(* IEC 61131-3 sources: plc-st-coding-agent/progress/evidence/f14_v13_self_20261113/jobs/diagnostic_deepseek-v4pro, 15 files *)

(* ---- public-easy-01.candidate_01.st ---- *)
(* ENGINEERING_CONTRACT
Independent retained outputs, all reset by finishedButton:
- Pump_Motor: set when bottleSensor TRUE, holds until finishedButton.
- Filling_Valve: set when cleaningConfirmButton TRUE, holds until finishedButton.
- Capping_Machine: set when fillingConfirmButton TRUE, holds until finishedButton.
- Packing_Machine: set when cappingConfirmButton TRUE, holds until finishedButton.
- Completion_Light: set when packingConfirmButton TRUE, reset by finishedButton.
Same-scan priority: finishedButton reset first, then trigger evaluations.
*)
(* CONTRACT_RULES [{"kind":"hold_until_reset","output":"Pump_Motor","set_input":"bottleSensor","reset_input":"finishedButton"},{"kind":"hold_until_reset","output":"Filling_Valve","set_input":"cleaningConfirmButton","reset_input":"finishedButton"},{"kind":"hold_until_reset","output":"Capping_Machine","set_input":"fillingConfirmButton","reset_input":"finishedButton"},{"kind":"hold_until_reset","output":"Packing_Machine","set_input":"cappingConfirmButton","reset_input":"finishedButton"},{"kind":"hold_until_reset","output":"Completion_Light","set_input":"packingConfirmButton","reset_input":"finishedButton"}] *)

FUNCTION_BLOCK FillingLineControl
VAR_INPUT
    bottleSensor : BOOL;
    cleaningConfirmButton : BOOL;
    fillingConfirmButton : BOOL;
    cappingConfirmButton : BOOL;
    packingConfirmButton : BOOL;
    finishedButton : BOOL;
END_VAR
VAR_OUTPUT
    Pump_Motor : BOOL;
    Filling_Valve : BOOL;
    Capping_Machine : BOOL;
    Packing_Machine : BOOL;
    Completion_Light : BOOL;
END_VAR
VAR
END_VAR

IF finishedButton THEN
    Pump_Motor := FALSE;
    Filling_Valve := FALSE;
    Capping_Machine := FALSE;
    Packing_Machine := FALSE;
    Completion_Light := FALSE;
ELSE
    IF bottleSensor THEN
        Pump_Motor := TRUE;
    END_IF;

    IF cleaningConfirmButton THEN
        Filling_Valve := TRUE;
    END_IF;

    IF fillingConfirmButton THEN
        Capping_Machine := TRUE;
    END_IF;

    IF cappingConfirmButton THEN
        Packing_Machine := TRUE;
    END_IF;

    IF packingConfirmButton THEN
        Completion_Light := TRUE;
    END_IF;
END_IF;

END_FUNCTION_BLOCK

(* ---- public-easy-01.candidate_02.st ---- *)
(* ENGINEERING_CONTRACT
Independent retained outputs, all reset by finishedButton:
- Pump_Motor: set when bottleSensor TRUE, holds until finishedButton.
- Filling_Valve: set when cleaningConfirmButton TRUE, holds until finishedButton.
- Capping_Machine: set when fillingConfirmButton TRUE, holds until finishedButton.
- Packing_Machine: set when cappingConfirmButton TRUE and Capping_Machine active, holds until finishedButton.
- Completion_Light: set when packingConfirmButton TRUE and Packing_Machine active, reset by finishedButton.
Same-scan priority: finishedButton reset first, then trigger evaluations.
*)
(* CONTRACT_RULES [{"kind":"hold_until_reset","output":"Pump_Motor","set_input":"bottleSensor","reset_input":"finishedButton"},{"kind":"hold_until_reset","output":"Filling_Valve","set_input":"cleaningConfirmButton","reset_input":"finishedButton"},{"kind":"hold_until_reset","output":"Capping_Machine","set_input":"fillingConfirmButton","reset_input":"finishedButton"}] *)

FUNCTION_BLOCK FillingLineControl
VAR_INPUT
    bottleSensor : BOOL;
    cleaningConfirmButton : BOOL;
    fillingConfirmButton : BOOL;
    cappingConfirmButton : BOOL;
    packingConfirmButton : BOOL;
    finishedButton : BOOL;
END_VAR
VAR_OUTPUT
    Pump_Motor : BOOL;
    Filling_Valve : BOOL;
    Capping_Machine : BOOL;
    Packing_Machine : BOOL;
    Completion_Light : BOOL;
END_VAR
VAR
END_VAR

IF finishedButton THEN
    Pump_Motor := FALSE;
    Filling_Valve := FALSE;
    Capping_Machine := FALSE;
    Packing_Machine := FALSE;
    Completion_Light := FALSE;
ELSE
    IF bottleSensor THEN
        Pump_Motor := TRUE;
    END_IF;

    IF cleaningConfirmButton THEN
        Filling_Valve := TRUE;
    END_IF;

    IF fillingConfirmButton THEN
        Capping_Machine := TRUE;
    END_IF;

    IF cappingConfirmButton AND Capping_Machine THEN
        Packing_Machine := TRUE;
    END_IF;

    IF packingConfirmButton AND Packing_Machine THEN
        Completion_Light := TRUE;
    END_IF;
END_IF;

END_FUNCTION_BLOCK

(* ---- public-easy-01.candidate_03.st ---- *)
(* ENGINEERING_CONTRACT
Independent retained outputs, all reset by finishedButton:
- Pump_Motor: set when bottleSensor TRUE, holds until finishedButton.
- Filling_Valve: set when cleaningConfirmButton TRUE, holds until finishedButton.
- Capping_Machine: set when fillingConfirmButton TRUE, holds until finishedButton.
- Packing_Machine: set when cappingConfirmButton TRUE and Capping_Machine active, holds until finishedButton.
- Completion_Light: set when packingConfirmButton TRUE and Packing_Machine active, reset by finishedButton.
Same-scan priority: finishedButton reset first, then trigger evaluations.
*)
(* CONTRACT_RULES [{"kind":"hold_until_reset","output":"Pump_Motor","set_input":"bottleSensor","reset_input":"finishedButton"},{"kind":"hold_until_reset","output":"Filling_Valve","set_input":"cleaningConfirmButton","reset_input":"finishedButton"},{"kind":"hold_until_reset","output":"Capping_Machine","set_input":"fillingConfirmButton","reset_input":"finishedButton"}] *)

FUNCTION_BLOCK FillingLineControl
VAR_INPUT
    bottleSensor : BOOL;
    cleaningConfirmButton : BOOL;
    fillingConfirmButton : BOOL;
    cappingConfirmButton : BOOL;
    packingConfirmButton : BOOL;
    finishedButton : BOOL;
END_VAR
VAR_OUTPUT
    Pump_Motor : BOOL;
    Filling_Valve : BOOL;
    Capping_Machine : BOOL;
    Packing_Machine : BOOL;
    Completion_Light : BOOL;
END_VAR
VAR
    local_PumpPrev : BOOL;
    local_FillingPrev : BOOL;
    local_CappingPrev : BOOL;
    local_PackingPrev : BOOL;
END_VAR

local_PumpPrev := Pump_Motor;
local_FillingPrev := Filling_Valve;
local_CappingPrev := Capping_Machine;
local_PackingPrev := Packing_Machine;

IF finishedButton THEN
    Pump_Motor := FALSE;
    Filling_Valve := FALSE;
    Capping_Machine := FALSE;
    Packing_Machine := FALSE;
    Completion_Light := FALSE;
ELSE
    IF bottleSensor THEN
        Pump_Motor := TRUE;
    END_IF;

    IF cleaningConfirmButton AND local_PumpPrev THEN
        Filling_Valve := TRUE;
    END_IF;

    IF fillingConfirmButton AND local_FillingPrev THEN
        Capping_Machine := TRUE;
    END_IF;

    IF cappingConfirmButton AND local_CappingPrev THEN
        Packing_Machine := TRUE;
    END_IF;

    IF packingConfirmButton AND local_PackingPrev THEN
        Completion_Light := TRUE;
    END_IF;
END_IF;

END_FUNCTION_BLOCK

(* ---- public-easy-01.patch_base_01.st ---- *)
(* ENGINEERING_CONTRACT
Outputs by state (state is persistent across scans):
- Pump_Motor: ON in CLEANING; starts when bottleSensor TRUE from IDLE; OFF on cleaningConfirmButton. Retained while CLEANING, even if bottleSensor falls (PUB001/PUB002).
- Filling_Valve: ON in FILLING; starts on cleaningConfirmButton in CLEANING; OFF on fillingConfirmButton (PUB002/PUB003).
- Capping_Machine: ON in CAPPING; starts on fillingConfirmButton in FILLING; OFF on cappingConfirmButton (PUB003/PUB004).
- Packing_Machine: ON in PACKING; starts on cappingConfirmButton in CAPPING; OFF on packingConfirmButton (PUB004/PUB005).
- Completion_Light: ON in COMPLETE; starts on packingConfirmButton in PACKING; reset by finishedButton (PUB005/PUB006/PUB007).
Same-scan priority: one state transition per call via ELSIF chain; outputs are assigned after transition using final state.
Buttons are treated as level-sensitive; pulse width/protocol unspecified.
*)
(* CONTRACT_RULES [] *)

FUNCTION_BLOCK FillingLineControl
VAR_INPUT
    bottleSensor: BOOL;
    cleaningConfirmButton: BOOL;
    fillingConfirmButton: BOOL;
    cappingConfirmButton: BOOL;
    packingConfirmButton: BOOL;
    finishedButton: BOOL;
END_VAR
VAR_OUTPUT
    Pump_Motor: BOOL;
    Filling_Valve: BOOL;
    Capping_Machine: BOOL;
    Packing_Machine: BOOL;
    Completion_Light: BOOL;
END_VAR
VAR
    step: INT := 0; (* 0=IDLE, 1=CLEANING, 2=FILLING, 3=CAPPING, 4=PACKING, 5=COMPLETE *)
    bottleTrig: R_TRIG;
END_VAR

(* State transitions: at most one per scan *)
bottleTrig(CLK := bottleSensor);

IF step = 0 THEN
    IF bottleTrig.Q THEN
        step := 1;
    END_IF;
ELSIF step = 1 THEN
    IF cleaningConfirmButton THEN
        step := 2;
    END_IF;
ELSIF step = 2 THEN
    IF fillingConfirmButton THEN
        step := 3;
    END_IF;
ELSIF step = 3 THEN
    IF cappingConfirmButton THEN
        step := 4;
    END_IF;
ELSIF step = 4 THEN
    IF packingConfirmButton THEN
        step := 5;
    END_IF;
ELSIF step = 5 THEN
    IF finishedButton THEN
        step := 0;
    END_IF;
END_IF;

(* Output mapping based on final state *)
CASE step OF
    0:
        Pump_Motor := FALSE;
        Filling_Valve := FALSE;
        Capping_Machine := FALSE;
        Packing_Machine := FALSE;
        Completion_Light := FALSE;

    1:
        Pump_Motor := TRUE;
        Filling_Valve := FALSE;
        Capping_Machine := FALSE;
        Packing_Machine := FALSE;
        Completion_Light := FALSE;

    2:
        Pump_Motor := FALSE;
        Filling_Valve := TRUE;
        Capping_Machine := FALSE;
        Packing_Machine := FALSE;
        Completion_Light := FALSE;

    3:
        Pump_Motor := FALSE;
        Filling_Valve := FALSE;
        Capping_Machine := TRUE;
        Packing_Machine := FALSE;
        Completion_Light := FALSE;

    4:
        Pump_Motor := FALSE;
        Filling_Valve := FALSE;
        Capping_Machine := FALSE;
        Packing_Machine := TRUE;
        Completion_Light := FALSE;

    5:
        Pump_Motor := FALSE;
        Filling_Valve := FALSE;
        Capping_Machine := FALSE;
        Packing_Machine := FALSE;
        Completion_Light := TRUE;

    ELSE
        Pump_Motor := FALSE;
        Filling_Valve := FALSE;
        Capping_Machine := FALSE;
        Packing_Machine := FALSE;
        Completion_Light := FALSE;
END_CASE;

END_FUNCTION_BLOCK

(* ---- public-easy-01.patch_base_02.st ---- *)
(* ENGINEERING_CONTRACT
Independent retained outputs, all reset by finishedButton:
- Pump_Motor: set when bottleSensor TRUE, holds until finishedButton.
- Filling_Valve: set when cleaningConfirmButton TRUE, holds until finishedButton.
- Capping_Machine: set when fillingConfirmButton TRUE, holds until finishedButton.
- Packing_Machine: set when cappingConfirmButton TRUE, holds until finishedButton.
- Completion_Light: set when packingConfirmButton TRUE, reset by finishedButton.
Same-scan priority: finishedButton reset first, then trigger evaluations.
*)
(* CONTRACT_RULES [{"kind":"hold_until_reset","output":"Pump_Motor","set_input":"bottleSensor","reset_input":"finishedButton"},{"kind":"hold_until_reset","output":"Filling_Valve","set_input":"cleaningConfirmButton","reset_input":"finishedButton"},{"kind":"hold_until_reset","output":"Capping_Machine","set_input":"fillingConfirmButton","reset_input":"finishedButton"},{"kind":"hold_until_reset","output":"Packing_Machine","set_input":"cappingConfirmButton","reset_input":"finishedButton"},{"kind":"hold_until_reset","output":"Completion_Light","set_input":"packingConfirmButton","reset_input":"finishedButton"}] *)

FUNCTION_BLOCK FillingLineControl
VAR_INPUT
    bottleSensor : BOOL;
    cleaningConfirmButton : BOOL;
    fillingConfirmButton : BOOL;
    cappingConfirmButton : BOOL;
    packingConfirmButton : BOOL;
    finishedButton : BOOL;
END_VAR
VAR_OUTPUT
    Pump_Motor : BOOL;
    Filling_Valve : BOOL;
    Capping_Machine : BOOL;
    Packing_Machine : BOOL;
    Completion_Light : BOOL;
END_VAR
VAR
END_VAR

IF finishedButton THEN
    Pump_Motor := FALSE;
    Filling_Valve := FALSE;
    Capping_Machine := FALSE;
    Packing_Machine := FALSE;
    Completion_Light := FALSE;
ELSE
    IF bottleSensor THEN
        Pump_Motor := TRUE;
    END_IF;

    IF cleaningConfirmButton THEN
        Filling_Valve := TRUE;
    END_IF;

    IF fillingConfirmButton THEN
        Capping_Machine := TRUE;
    END_IF;

    IF cappingConfirmButton THEN
        Packing_Machine := TRUE;
    END_IF;

    IF packingConfirmButton THEN
        Completion_Light := TRUE;
    END_IF;
END_IF;

END_FUNCTION_BLOCK

(* ---- public-easy-01.patch_base_03.st ---- *)
(* ENGINEERING_CONTRACT
Independent retained outputs, all reset by finishedButton:
- Pump_Motor: set when bottleSensor TRUE, holds until finishedButton.
- Filling_Valve: set when cleaningConfirmButton TRUE, holds until finishedButton.
- Capping_Machine: set when fillingConfirmButton TRUE, holds until finishedButton.
- Packing_Machine: set when cappingConfirmButton TRUE and Capping_Machine active, holds until finishedButton.
- Completion_Light: set when packingConfirmButton TRUE and Packing_Machine active, reset by finishedButton.
Same-scan priority: finishedButton reset first, then trigger evaluations.
*)
(* CONTRACT_RULES [{"kind":"hold_until_reset","output":"Pump_Motor","set_input":"bottleSensor","reset_input":"finishedButton"},{"kind":"hold_until_reset","output":"Filling_Valve","set_input":"cleaningConfirmButton","reset_input":"finishedButton"},{"kind":"hold_until_reset","output":"Capping_Machine","set_input":"fillingConfirmButton","reset_input":"finishedButton"}] *)

FUNCTION_BLOCK FillingLineControl
VAR_INPUT
    bottleSensor : BOOL;
    cleaningConfirmButton : BOOL;
    fillingConfirmButton : BOOL;
    cappingConfirmButton : BOOL;
    packingConfirmButton : BOOL;
    finishedButton : BOOL;
END_VAR
VAR_OUTPUT
    Pump_Motor : BOOL;
    Filling_Valve : BOOL;
    Capping_Machine : BOOL;
    Packing_Machine : BOOL;
    Completion_Light : BOOL;
END_VAR
VAR
END_VAR

IF finishedButton THEN
    Pump_Motor := FALSE;
    Filling_Valve := FALSE;
    Capping_Machine := FALSE;
    Packing_Machine := FALSE;
    Completion_Light := FALSE;
ELSE
    IF bottleSensor THEN
        Pump_Motor := TRUE;
    END_IF;

    IF cleaningConfirmButton THEN
        Filling_Valve := TRUE;
    END_IF;

    IF fillingConfirmButton THEN
        Capping_Machine := TRUE;
    END_IF;

    IF cappingConfirmButton AND Capping_Machine THEN
        Packing_Machine := TRUE;
    END_IF;

    IF packingConfirmButton AND Packing_Machine THEN
        Completion_Light := TRUE;
    END_IF;
END_IF;

END_FUNCTION_BLOCK

(* ---- public-easy-01.raw_candidate_01.st ---- *)
(* ENGINEERING_CONTRACT
Independent retained outputs, all reset by finishedButton:
- Pump_Motor: set when bottleSensor TRUE, holds until finishedButton.
- Filling_Valve: set when cleaningConfirmButton TRUE, holds until finishedButton.
- Capping_Machine: set when fillingConfirmButton TRUE, holds until finishedButton.
- Packing_Machine: set when cappingConfirmButton TRUE, holds until finishedButton.
- Completion_Light: set when packingConfirmButton TRUE, reset by finishedButton.
Same-scan priority: finishedButton reset first, then trigger evaluations.
*)
(* CONTRACT_RULES [{"kind":"hold_until_reset","output":"Pump_Motor","set_input":"bottleSensor","reset_input":"finishedButton"},{"kind":"hold_until_reset","output":"Filling_Valve","set_input":"cleaningConfirmButton","reset_input":"finishedButton"},{"kind":"hold_until_reset","output":"Capping_Machine","set_input":"fillingConfirmButton","reset_input":"finishedButton"},{"kind":"hold_until_reset","output":"Packing_Machine","set_input":"cappingConfirmButton","reset_input":"finishedButton"},{"kind":"hold_until_reset","output":"Completion_Light","set_input":"packingConfirmButton","reset_input":"finishedButton"}] *)

FUNCTION_BLOCK FillingLineControl
VAR_INPUT
    bottleSensor : BOOL;
    cleaningConfirmButton : BOOL;
    fillingConfirmButton : BOOL;
    cappingConfirmButton : BOOL;
    packingConfirmButton : BOOL;
    finishedButton : BOOL;
END_VAR
VAR_OUTPUT
    Pump_Motor : BOOL;
    Filling_Valve : BOOL;
    Capping_Machine : BOOL;
    Packing_Machine : BOOL;
    Completion_Light : BOOL;
END_VAR
VAR
END_VAR

IF finishedButton THEN
    Pump_Motor := FALSE;
    Filling_Valve := FALSE;
    Capping_Machine := FALSE;
    Packing_Machine := FALSE;
    Completion_Light := FALSE;
ELSE
    IF bottleSensor THEN
        Pump_Motor := TRUE;
    END_IF;

    IF cleaningConfirmButton THEN
        Filling_Valve := TRUE;
    END_IF;

    IF fillingConfirmButton THEN
        Capping_Machine := TRUE;
    END_IF;

    IF cappingConfirmButton THEN
        Packing_Machine := TRUE;
    END_IF;

    IF packingConfirmButton THEN
        Completion_Light := TRUE;
    END_IF;
END_IF;

END_FUNCTION_BLOCK

(* ---- public-easy-01.raw_candidate_02.st ---- *)
(* ENGINEERING_CONTRACT
Independent retained outputs, all reset by finishedButton:
- Pump_Motor: set when bottleSensor TRUE, holds until finishedButton.
- Filling_Valve: set when cleaningConfirmButton TRUE, holds until finishedButton.
- Capping_Machine: set when fillingConfirmButton TRUE, holds until finishedButton.
- Packing_Machine: set when cappingConfirmButton TRUE and Capping_Machine active, holds until finishedButton.
- Completion_Light: set when packingConfirmButton TRUE and Packing_Machine active, reset by finishedButton.
Same-scan priority: finishedButton reset first, then trigger evaluations.
*)
(* CONTRACT_RULES [{"kind":"hold_until_reset","output":"Pump_Motor","set_input":"bottleSensor","reset_input":"finishedButton"},{"kind":"hold_until_reset","output":"Filling_Valve","set_input":"cleaningConfirmButton","reset_input":"finishedButton"},{"kind":"hold_until_reset","output":"Capping_Machine","set_input":"fillingConfirmButton","reset_input":"finishedButton"}] *)

FUNCTION_BLOCK FillingLineControl
VAR_INPUT
    bottleSensor : BOOL;
    cleaningConfirmButton : BOOL;
    fillingConfirmButton : BOOL;
    cappingConfirmButton : BOOL;
    packingConfirmButton : BOOL;
    finishedButton : BOOL;
END_VAR
VAR_OUTPUT
    Pump_Motor : BOOL;
    Filling_Valve : BOOL;
    Capping_Machine : BOOL;
    Packing_Machine : BOOL;
    Completion_Light : BOOL;
END_VAR
VAR
END_VAR

IF finishedButton THEN
    Pump_Motor := FALSE;
    Filling_Valve := FALSE;
    Capping_Machine := FALSE;
    Packing_Machine := FALSE;
    Completion_Light := FALSE;
ELSE
    IF bottleSensor THEN
        Pump_Motor := TRUE;
    END_IF;

    IF cleaningConfirmButton THEN
        Filling_Valve := TRUE;
    END_IF;

    IF fillingConfirmButton THEN
        Capping_Machine := TRUE;
    END_IF;

    IF cappingConfirmButton AND Capping_Machine THEN
        Packing_Machine := TRUE;
    END_IF;

    IF packingConfirmButton AND Packing_Machine THEN
        Completion_Light := TRUE;
    END_IF;
END_IF;

END_FUNCTION_BLOCK

(* ---- public-easy-01.raw_candidate_03.st ---- *)
(* ENGINEERING_CONTRACT
Independent retained outputs, all reset by finishedButton:
- Pump_Motor: set when bottleSensor TRUE, holds until finishedButton.
- Filling_Valve: set when cleaningConfirmButton TRUE, holds until finishedButton.
- Capping_Machine: set when fillingConfirmButton TRUE, holds until finishedButton.
- Packing_Machine: set when cappingConfirmButton TRUE and Capping_Machine active, holds until finishedButton.
- Completion_Light: set when packingConfirmButton TRUE and Packing_Machine active, reset by finishedButton.
Same-scan priority: finishedButton reset first, then trigger evaluations.
*)
(* CONTRACT_RULES [{"kind":"hold_until_reset","output":"Pump_Motor","set_input":"bottleSensor","reset_input":"finishedButton"},{"kind":"hold_until_reset","output":"Filling_Valve","set_input":"cleaningConfirmButton","reset_input":"finishedButton"},{"kind":"hold_until_reset","output":"Capping_Machine","set_input":"fillingConfirmButton","reset_input":"finishedButton"}] *)

FUNCTION_BLOCK FillingLineControl
VAR_INPUT
    bottleSensor : BOOL;
    cleaningConfirmButton : BOOL;
    fillingConfirmButton : BOOL;
    cappingConfirmButton : BOOL;
    packingConfirmButton : BOOL;
    finishedButton : BOOL;
END_VAR
VAR_OUTPUT
    Pump_Motor : BOOL;
    Filling_Valve : BOOL;
    Capping_Machine : BOOL;
    Packing_Machine : BOOL;
    Completion_Light : BOOL;
END_VAR
VAR
    local_PumpPrev : BOOL;
    local_FillingPrev : BOOL;
    local_CappingPrev : BOOL;
    local_PackingPrev : BOOL;
END_VAR

local_PumpPrev := Pump_Motor;
local_FillingPrev := Filling_Valve;
local_CappingPrev := Capping_Machine;
local_PackingPrev := Packing_Machine;

IF finishedButton THEN
    Pump_Motor := FALSE;
    Filling_Valve := FALSE;
    Capping_Machine := FALSE;
    Packing_Machine := FALSE;
    Completion_Light := FALSE;
ELSE
    IF bottleSensor THEN
        Pump_Motor := TRUE;
    END_IF;

    IF cleaningConfirmButton AND local_PumpPrev THEN
        Filling_Valve := TRUE;
    END_IF;

    IF fillingConfirmButton AND local_FillingPrev THEN
        Capping_Machine := TRUE;
    END_IF;

    IF cappingConfirmButton AND local_CappingPrev THEN
        Packing_Machine := TRUE;
    END_IF;

    IF packingConfirmButton AND local_PackingPrev THEN
        Completion_Light := TRUE;
    END_IF;
END_IF;

END_FUNCTION_BLOCK

(* ---- public-hard-04.candidate_01.st ---- *)
(* ENGINEERING_CONTRACT
   elementCount DINT: retained process value; 0 after reset, +1 successful enqueue, -1 successful dequeue, held otherwise; range 0..capacity.
   status WORD: overwritten every invocation; 0 idle/reset/success, 16#8002 rejected full enqueue, 16#8001 rejected empty dequeue; reset priority sets 0.
   queue state: first invocation empty; reset priority clears head/tail/count; enqueue writes at tail, dequeue reads head; circular indices low..high.
   edge triggers: R_TRIG consumed every scan; reset priority ignores edge requests; simultaneous enqueue+dequeue unspecified -> no-op.
   units/boundaries: capacity positive DINT derived each scan from LOWER_BOUND/UPPER_BOUND of the supplied array; first element index may be nonzero.
*)
(* CONTRACT_RULES [] *)
FUNCTION_BLOCK FIFO
VAR_INPUT
    enqueue : BOOL;
    dequeue : BOOL;
    reset : BOOL;
END_VAR
VAR_OUTPUT
    elementCount : DINT;
    status : WORD;
END_VAR
VAR_IN_OUT
    item : VARIANT;
    buffer : VARIANT;
END_VAR
VAR
    local_rEnq : R_TRIG;
    local_rDeq : R_TRIG;
    local_enqEdge : BOOL;
    local_deqEdge : BOOL;

    local_low : DINT;
    local_high : DINT;
    local_capacity : DINT;
    local_count : DINT := 0;
    local_head : DINT := 0;
    local_tail : DINT := 0;
END_VAR

local_rEnq(CLK := enqueue);
local_enqEdge := local_rEnq.Q;
local_rDeq(CLK := dequeue);
local_deqEdge := local_rDeq.Q;

status := 16#0000;

local_low := LOWER_BOUND(buffer, 1);
local_high := UPPER_BOUND(buffer, 1);
local_capacity := local_high - local_low + 1;
IF local_capacity < 1 THEN
    local_capacity := 1;
END_IF;

IF local_count = 0 THEN
    local_head := local_low;
    local_tail := local_low;
END_IF;

IF reset THEN
    local_count := 0;
    local_head := local_low;
    local_tail := local_low;
    status := 16#0000;
ELSE
    IF local_enqEdge AND NOT local_deqEdge THEN
        IF local_count < local_capacity THEN
            buffer[local_tail] := item;
            local_tail := local_tail + 1;
            IF local_tail > local_high THEN
                local_tail := local_low;
            END_IF;
            local_count := local_count + 1;
            status := 16#0000;
        ELSE
            status := 16#8002;
        END_IF;
    ELSIF local_deqEdge AND NOT local_enqEdge THEN
        IF local_count > 0 THEN
            item := buffer[local_head];
            local_head := local_head + 1;
            IF local_head > local_high THEN
                local_head := local_low;
            END_IF;
            local_count := local_count - 1;
            status := 16#0000;
        ELSE
            status := 16#8001;
        END_IF;
    END_IF;
END_IF;

elementCount := local_count;

(* ---- public-hard-04.candidate_02.st ---- *)
(* ENGINEERING_CONTRACT
   elementCount DINT: retained process value; 0 after reset, +1 successful enqueue, -1 successful dequeue, held otherwise; range 0..capacity.
   status WORD: overwritten every invocation; 0 idle/reset/success, 16#8002 rejected full enqueue, 16#8001 rejected empty dequeue; reset priority sets 0.
   queue state: first invocation empty; reset priority clears head/tail/count; enqueue writes at tail, dequeue reads head; circular indices low..high.
   edge triggers: R_TRIG consumed every scan; reset priority ignores edge requests; simultaneous enqueue+dequeue unspecified -> no-op.
   units/boundaries: capacity positive DINT derived each scan from LOWER_BOUND/UPPER_BOUND of the supplied array; first element index may be nonzero.
*)
(* CONTRACT_RULES [] *)
FUNCTION_BLOCK FIFO
VAR_INPUT
    enqueue : BOOL;
    dequeue : BOOL;
    reset : BOOL;
END_VAR
VAR_OUTPUT
    elementCount : DINT;
    status : WORD;
END_VAR
VAR_IN_OUT
    item : VARIANT;
    buffer : VARIANT;
END_VAR
VAR
    local_rEnq : R_TRIG;
    local_rDeq : R_TRIG;
    local_enqEdge : BOOL;
    local_deqEdge : BOOL;

    local_low : DINT;
    local_high : DINT;
    local_capacity : DINT;
    local_count : DINT := 0;
    local_head : DINT := 0;
    local_tail : DINT := 0;
END_VAR

local_rEnq(CLK := enqueue);
local_enqEdge := local_rEnq.Q;
local_rDeq(CLK := dequeue);
local_deqEdge := local_rDeq.Q;

status := 16#0000;

local_low := LOWER_BOUND(buffer, 1);
local_high := UPPER_BOUND(buffer, 1);
local_capacity := local_high - local_low + 1;
IF local_capacity < 1 THEN
    local_capacity := 1;
END_IF;

IF local_count = 0 THEN
    local_head := local_low;
    local_tail := local_low;
END_IF;

IF reset THEN
    local_count := 0;
    local_head := local_low;
    local_tail := local_low;
    status := 16#0000;
ELSE
    IF local_enqEdge AND NOT local_deqEdge THEN
        IF local_count < local_capacity THEN
            buffer[local_tail] := item;
            local_tail := local_tail + 1;
            IF local_tail > local_high THEN
                local_tail := local_low;
            END_IF;
            local_count := local_count + 1;
            status := 16#0000;
        ELSE
            status := 16#8002;
        END_IF;
    ELSIF local_deqEdge AND NOT local_enqEdge THEN
        IF local_count > 0 THEN
            item := buffer[local_head];
            local_head := local_head + 1;
            IF local_head > local_high THEN
                local_head := local_low;
            END_IF;
            local_count := local_count - 1;
            status := 16#0000;
        ELSE
            status := 16#8001;
        END_IF;
    END_IF;
END_IF;

elementCount := local_count;

END_FUNCTION_BLOCK

(* ---- public-hard-04.patch_base_01.st ---- *)
(* ENGINEERING_CONTRACT
   elementCount DINT: retained process value; 0 after reset, +1 successful enqueue, -1 successful dequeue, held otherwise; range 0..capacity.
   status WORD: overwritten every invocation; 0 idle/reset/success, 16#8002 rejected full enqueue, 16#8001 rejected empty dequeue; reset priority sets 0.
   queue state: first invocation empty; reset priority clears head/tail/count; enqueue writes at tail, dequeue reads head; indices 0..capacity-1.
   edge triggers: R_TRIG consumed every scan; reset priority ignores edge requests; simultaneous enqueue+dequeue unspecified -> no-op.
   units/boundaries: capacity positive DINT derived once from buffer size / item element size; element copied byte-wise from item address.
*)
(* CONTRACT_RULES [] *)
FUNCTION_BLOCK FIFO
VAR_INPUT
    enqueue : BOOL;
    dequeue : BOOL;
    reset : BOOL;
END_VAR
VAR_OUTPUT
    elementCount : DINT;
    status : WORD;
END_VAR
VAR_IN_OUT
    item : VARIANT;
    buffer : VARIANT;
END_VAR
VAR
    local_rEnq : R_TRIG;
    local_rDeq : R_TRIG;
    local_enqEdge : BOOL;
    local_deqEdge : BOOL;

    local_associated : BOOL := FALSE;
    local_pBufferBase : POINTER TO BYTE;
    local_pItemBase : POINTER TO BYTE;
    local_elemSize : DINT := 1;
    local_capacity : DINT := 1;

    local_count : DINT := 0;
    local_head : DINT := 0;
    local_tail : DINT := 0;

    local_bufInfo : __SYSTEM.VAR_INFO;
    local_itemInfo : __SYSTEM.VAR_INFO;

    local_pSrc : POINTER TO BYTE;
    local_pDst : POINTER TO BYTE;
    local_i : DINT;
END_VAR

(* Consume rising edges every scan so reset cannot create ghost operations later. *)
local_rEnq(CLK := enqueue);
local_enqEdge := local_rEnq.Q;
local_rDeq(CLK := dequeue);
local_deqEdge := local_rDeq.Q;

status := 16#0000;

(* One-time association of buffer and element storage, using the first invocation. *)
IF NOT local_associated THEN
    local_bufInfo := __VARINFO(buffer);
    local_itemInfo := __VARINFO(item);

    local_elemSize := local_itemInfo.diSize;
    IF local_elemSize <= 0 THEN
        local_elemSize := 1;
    END_IF;

    local_capacity := local_bufInfo.diSize / local_elemSize;
    IF local_capacity < 1 THEN
        local_capacity := 1;
    END_IF;

    local_pBufferBase := local_bufInfo.pvAddress;
    local_pItemBase := local_itemInfo.pvAddress;
    local_associated := TRUE;
END_IF;

IF reset THEN
    (* Reset has priority over all operations; stored values remain untouched. *)
    local_count := 0;
    local_head := 0;
    local_tail := 0;
    status := 16#0000;
ELSE
    IF local_enqEdge AND NOT local_deqEdge THEN
        IF local_count < local_capacity THEN
            (* Copy current item value into tail slot. *)
            local_pSrc := local_pItemBase;
            local_pDst := local_pBufferBase + (local_tail * local_elemSize);

            FOR local_i := 0 TO local_elemSize - 1 DO
                local_pDst^ := local_pSrc^;
                local_pSrc := local_pSrc + 1;
                local_pDst := local_pDst + 1;
            END_FOR;

            local_tail := (local_tail + 1) MOD local_capacity;
            local_count := local_count + 1;
            status := 16#0000;
        ELSE
            status := 16#8002; (* enqueue rejected: full *)
        END_IF;
    ELSIF local_deqEdge AND NOT local_enqEdge THEN
        IF local_count > 0 THEN
            (* Copy head element back to item. *)
            local_pSrc := local_pBufferBase + (local_head * local_elemSize);
            local_pDst := local_pItemBase;

            FOR local_i := 0 TO local_elemSize - 1 DO
                local_pDst^ := local_pSrc^;
                local_pSrc := local_pSrc + 1;
                local_pDst := local_pDst + 1;
            END_FOR;

            local_head := (local_head + 1) MOD local_capacity;
            local_count := local_count - 1;
            status := 16#0000;
        ELSE
            status := 16#8001; (* dequeue rejected: empty *)
        END_IF;
    END_IF;
END_IF;

elementCount := local_count;

(* ---- public-hard-04.patch_base_02.st ---- *)
(* ENGINEERING_CONTRACT
   elementCount DINT: retained process value; 0 after reset, +1 successful enqueue, -1 successful dequeue, held otherwise; range 0..capacity.
   status WORD: overwritten every invocation; 0 idle/reset/success, 16#8002 rejected full enqueue, 16#8001 rejected empty dequeue; reset priority sets 0.
   queue state: first invocation empty; reset priority clears head/tail/count; enqueue writes at tail, dequeue reads head; circular indices low..high.
   edge triggers: R_TRIG consumed every scan; reset priority ignores edge requests; simultaneous enqueue+dequeue unspecified -> no-op.
   units/boundaries: capacity positive DINT derived each scan from LOWER_BOUND/UPPER_BOUND of the supplied array; first element index may be nonzero.
*)
(* CONTRACT_RULES [] *)
FUNCTION_BLOCK FIFO
VAR_INPUT
    enqueue : BOOL;
    dequeue : BOOL;
    reset : BOOL;
END_VAR
VAR_OUTPUT
    elementCount : DINT;
    status : WORD;
END_VAR
VAR_IN_OUT
    item : VARIANT;
    buffer : VARIANT;
END_VAR
VAR
    local_rEnq : R_TRIG;
    local_rDeq : R_TRIG;
    local_enqEdge : BOOL;
    local_deqEdge : BOOL;

    local_low : DINT;
    local_high : DINT;
    local_capacity : DINT;
    local_count : DINT := 0;
    local_head : DINT := 0;
    local_tail : DINT := 0;
END_VAR

local_rEnq(CLK := enqueue);
local_enqEdge := local_rEnq.Q;
local_rDeq(CLK := dequeue);
local_deqEdge := local_rDeq.Q;

status := 16#0000;

local_low := LOWER_BOUND(buffer, 1);
local_high := UPPER_BOUND(buffer, 1);
local_capacity := local_high - local_low + 1;
IF local_capacity < 1 THEN
    local_capacity := 1;
END_IF;

IF local_count = 0 THEN
    local_head := local_low;
    local_tail := local_low;
END_IF;

IF reset THEN
    local_count := 0;
    local_head := local_low;
    local_tail := local_low;
    status := 16#0000;
ELSE
    IF local_enqEdge AND NOT local_deqEdge THEN
        IF local_count < local_capacity THEN
            buffer[local_tail] := item;
            local_tail := local_tail + 1;
            IF local_tail > local_high THEN
                local_tail := local_low;
            END_IF;
            local_count := local_count + 1;
            status := 16#0000;
        ELSE
            status := 16#8002;
        END_IF;
    ELSIF local_deqEdge AND NOT local_enqEdge THEN
        IF local_count > 0 THEN
            item := buffer[local_head];
            local_head := local_head + 1;
            IF local_head > local_high THEN
                local_head := local_low;
            END_IF;
            local_count := local_count - 1;
            status := 16#0000;
        ELSE
            status := 16#8001;
        END_IF;
    END_IF;
END_IF;

elementCount := local_count;

(* ---- public-hard-04.raw_candidate_01.st ---- *)
(* ENGINEERING_CONTRACT
   elementCount DINT: retained process value; 0 after reset, +1 successful enqueue, -1 successful dequeue, held otherwise; range 0..capacity.
   status WORD: overwritten every invocation; 0 idle/reset/success, 16#8002 rejected full enqueue, 16#8001 rejected empty dequeue; reset priority sets 0.
   queue state: first invocation empty; reset priority clears head/tail/count; enqueue writes at tail, dequeue reads head; circular indices low..high.
   edge triggers: R_TRIG consumed every scan; reset priority ignores edge requests; simultaneous enqueue+dequeue unspecified -> no-op.
   units/boundaries: capacity positive DINT derived each scan from LOWER_BOUND/UPPER_BOUND of the supplied array; first element index may be nonzero.
*)
(* CONTRACT_RULES [] *)
FUNCTION_BLOCK FIFO
VAR_INPUT
    enqueue : BOOL;
    dequeue : BOOL;
    reset : BOOL;
END_VAR
VAR_OUTPUT
    elementCount : DINT;
    status : WORD;
END_VAR
VAR_IN_OUT
    item : VARIANT;
    buffer : VARIANT;
END_VAR
VAR
    local_rEnq : R_TRIG;
    local_rDeq : R_TRIG;
    local_enqEdge : BOOL;
    local_deqEdge : BOOL;

    local_low : DINT;
    local_high : DINT;
    local_capacity : DINT;
    local_count : DINT := 0;
    local_head : DINT := 0;
    local_tail : DINT := 0;
END_VAR

local_rEnq(CLK := enqueue);
local_enqEdge := local_rEnq.Q;
local_rDeq(CLK := dequeue);
local_deqEdge := local_rDeq.Q;

status := 16#0000;

local_low := LOWER_BOUND(buffer, 1);
local_high := UPPER_BOUND(buffer, 1);
local_capacity := local_high - local_low + 1;
IF local_capacity < 1 THEN
    local_capacity := 1;
END_IF;

IF local_count = 0 THEN
    local_head := local_low;
    local_tail := local_low;
END_IF;

IF reset THEN
    local_count := 0;
    local_head := local_low;
    local_tail := local_low;
    status := 16#0000;
ELSE
    IF local_enqEdge AND NOT local_deqEdge THEN
        IF local_count < local_capacity THEN
            buffer[local_tail] := item;
            local_tail := local_tail + 1;
            IF local_tail > local_high THEN
                local_tail := local_low;
            END_IF;
            local_count := local_count + 1;
            status := 16#0000;
        ELSE
            status := 16#8002;
        END_IF;
    ELSIF local_deqEdge AND NOT local_enqEdge THEN
        IF local_count > 0 THEN
            item := buffer[local_head];
            local_head := local_head + 1;
            IF local_head > local_high THEN
                local_head := local_low;
            END_IF;
            local_count := local_count - 1;
            status := 16#0000;
        ELSE
            status := 16#8001;
        END_IF;
    END_IF;
END_IF;

elementCount := local_count;

(* ---- public-hard-04.raw_candidate_02.st ---- *)
(* ENGINEERING_CONTRACT
   elementCount DINT: retained process value; 0 after reset, +1 successful enqueue, -1 successful dequeue, held otherwise; range 0..capacity.
   status WORD: overwritten every invocation; 0 idle/reset/success, 16#8002 rejected full enqueue, 16#8001 rejected empty dequeue; reset priority sets 0.
   queue state: first invocation empty; reset priority clears head/tail/count; enqueue writes at tail, dequeue reads head; circular indices low..high.
   edge triggers: R_TRIG consumed every scan; reset priority ignores edge requests; simultaneous enqueue+dequeue unspecified -> no-op.
   units/boundaries: capacity positive DINT derived each scan from LOWER_BOUND/UPPER_BOUND of the supplied array; first element index may be nonzero.
*)
(* CONTRACT_RULES [] *)
FUNCTION_BLOCK FIFO
VAR_INPUT
    enqueue : BOOL;
    dequeue : BOOL;
    reset : BOOL;
END_VAR
VAR_OUTPUT
    elementCount : DINT;
    status : WORD;
END_VAR
VAR_IN_OUT
    item : VARIANT;
    buffer : VARIANT;
END_VAR
VAR
    local_rEnq : R_TRIG;
    local_rDeq : R_TRIG;
    local_enqEdge : BOOL;
    local_deqEdge : BOOL;

    local_low : DINT;
    local_high : DINT;
    local_capacity : DINT;
    local_count : DINT := 0;
    local_head : DINT := 0;
    local_tail : DINT := 0;
END_VAR

local_rEnq(CLK := enqueue);
local_enqEdge := local_rEnq.Q;
local_rDeq(CLK := dequeue);
local_deqEdge := local_rDeq.Q;

status := 16#0000;

local_low := LOWER_BOUND(buffer, 1);
local_high := UPPER_BOUND(buffer, 1);
local_capacity := local_high - local_low + 1;
IF local_capacity < 1 THEN
    local_capacity := 1;
END_IF;

IF local_count = 0 THEN
    local_head := local_low;
    local_tail := local_low;
END_IF;

IF reset THEN
    local_count := 0;
    local_head := local_low;
    local_tail := local_low;
    status := 16#0000;
ELSE
    IF local_enqEdge AND NOT local_deqEdge THEN
        IF local_count < local_capacity THEN
            buffer[local_tail] := item;
            local_tail := local_tail + 1;
            IF local_tail > local_high THEN
                local_tail := local_low;
            END_IF;
            local_count := local_count + 1;
            status := 16#0000;
        ELSE
            status := 16#8002;
        END_IF;
    ELSIF local_deqEdge AND NOT local_enqEdge THEN
        IF local_count > 0 THEN
            item := buffer[local_head];
            local_head := local_head + 1;
            IF local_head > local_high THEN
                local_head := local_low;
            END_IF;
            local_count := local_count - 1;
            status := 16#0000;
        ELSE
            status := 16#8001;
        END_IF;
    END_IF;
END_IF;

elementCount := local_count;

END_FUNCTION_BLOCK
